Staubli VAL3: trajItem.dtx

public num nFrameIndex
public num nToolIndex
public string sID
public num nMoveID
public pointItem pPointItem
  [0]
    pointRx pPointRx[2]
    jointRx jJointRx
    paraItem pParaItem
      [0]
        mdesc mMdesc
        num nMoveType
        num nActionIndex
        num nPercentage
        ifItem iIfItem
          [0]
            num nSigType[3]
            num nSigIndex[3]
            num nValue[3]
            bool bANDOR[2]
        num nDelay
        num nSigValue
        bool bSafePoint
    string sID
    bool bMarked
    pointRx pInter
